(* IEC 61131-3 sources: traffic-lights/PLC_TrafficLights/Class/HwControl (part 2) *)

      ret_code                := BUSY;

      StartTime               := ops.tAbsolute;
      AdditionalPostInitTime  := 0;
      sd_retval               := 0;

//**********************************************************************************************************************************************************
//** CALCULATE, SET AND DISTRIBUTE TASK TIMES                                                                                                             **
//**********************************************************************************************************************************************************

      for i:=0 to TASK_SELECT_COREMAX do

      //Calculate Tasksettings for each core
        CalculateTaskInfo(us_CoreSelect:=i$USINT, pTaskInfo:=#aTaskInfoCore[i]);

        //Special Core 0 has to be running in RtWork method (is needed because if we dont have the new interfaces we cannot move a function to first realtime pos later)
        //Always add Realtime and Cyclic for Core 0: Realtime of Core 0 does watchdog trigger and calls for Diasmaster
        //***********************************************************
        if aTaskInfoCore[i].us_CoreSelect = TASK_SELECT_CORE0 then

          //Rt Prescan
          //**********************************************************************************************************************************************

          //get objectinfo of HwControl object
          //maybe we have a derivation with configured realtime task --> we have to change the task time of the task to the correct setting
          sd_retval := To_TaskObjectControl.GetObjectInfo( thispointer := this, tasktype := OBJ_RT, objinfo := #s_objinfo);

          //Check if we have a configured tasktime
          if sd_retval <> 0 | s_objinfo.period = 0 then

            //No task configured --> use OS function to add the RT Task

            //Note: udPhase must always be TASK_SCAN. At RTK there was an error that using TASK_PRE and TASK_POST occurs an access-exception in the OS.
            //With TASK_SCAN the object/function will be added in the list at the end. (will be moved to first position later if needed)
            if OS_AddRtObject(udMode  := TASK_TIMED
                            , udTime  := aTaskInfoCore[i].ud_MyRtTaskTime_us OR 16#8000_0000
                            , udPhase := TASK_SCAN) = NIL then
              HWC_LogValue1(this,"@0160 (HWControl::Control::NewInst) OS_AddRtObject failed to add Realtime (Prescan) object for core 0x{0}",aTaskInfoCore[i].us_CoreSelect);
            end_if;
          else

            // User must have a derivation of the HWControl with a configured Realtime Task --> Change the task time of the existing realtime task
            if To_TaskObjectControl.ChangeObjectState(thispointer :=  this
                                                    , actioncmd   :=  ACTION_NEWTIME
                                                    , tasktype    :=  OBJ_RT
                                                    , debugobj    :=  0
                                                    , newtime     :=  aTaskInfoCore[i].ud_MyRtTaskTime_us OR 16#8000_0000
                                                    ) <> 0 then
              HWC_LogError(this,"@03E3 (HWControl::Control::NewInst) Failed to change the object state to set the correct realtime task settings.");
            end_if;
          end_if;

          //RT Postscan
          //**********************************************************************************************************************************************

          //Check for Rt-Debug State. Do not add the Rt func for postscan if RtDebug is activated (because postscan will be called from prescan in this case)

          if GetRtDebugState() = TRUE then
            //save thispointer of object in OS-function (leads to that the task is called from the Breakpoint handler from the OS so the user can debug and the Hwcontrol is still running (no watchdog error))
            if p_DebugAPI then
              SaveThisPointer( this, TASK_SELECT_CORE0 );
            else
              HWC_LogError(this,"@0167 (HWControl::Control::NewInst) Pointer p_DebugAPI is invalid. Rt-Debug is not supported");
            end_if;

            // Set RtPostScan off if RtDebug is used!
            if To_TaskObjectControl.ChangeObjectState(thispointer :=  #HWRtPostScan.ClassSvr$void
                                                    , actioncmd   :=  ACTION_SUSPEND
                                                    , tasktype    :=  OBJ_RT
                                                    , debugobj    :=  0
                                                    , newtime     :=  0
                                                    ) <> 0 then
              HWC_LogError(this,"@0161 (HWControl::Control::NewInst) Failed to change object state of HwRtPostscan object");
            end_if;

          else

            //We have to use the object of HwRtPostscan instead of using the function OS_AddRtObject due to problems with RTK-CPUs (e.g. CP212)
            //The problem is that, with a maintimer of 500µs, and a task time of 1ms it can happen that the realtime (prescan) and the postscan of this class
            //are not "synchronized", which means that they have a time gap of 500µs between each other which leads to problems (TimesliceError).
            //This is not a problem with Salamander CPUs (e.g CP111)

            // Synchronize calls of Rt & RtPostScan (same timebase)
            if To_TaskObjectControl.ChangeObjectState(thispointer :=  #HWRtPostScan.ClassSvr$void
                                                    , actioncmd   :=  ACTION_NEWTIME
                                                    , tasktype    :=  OBJ_RT
                                                    , debugobj    :=  0
                                                    , newtime     :=  aTaskInfoCore[i].ud_MyRtTaskTime_us OR 16#8000_0000
                                                    ) <> 0 then
              HWC_LogError(this,"@0161 (HWControl::Control::NewInst) Failed to change object state of HwRtPostscan object");
            end_if;

            //save NIL-Pointer to OS-function because only HwControl is allowed to use this function
            if p_DebugAPI then
              SaveThisPointer( NIL, TASK_SELECT_CORE0 );
            end_if;

            //rt-post scan is added - realtime is added
            sRtTaskControl.usCoresRtActive  += 1;

          end_if;

          //Cyclic Task
          //**********************************************************************************************************************************************

          //Note: OS_AddCyFunc can NOT be used!! On RTK-CPUs with emulated SRAM () it leads to a reboot of the CPU if the SRAM is accessed from a function that is added via OS_AddCyFunc (or OS_AddRtFunc).
//          if OS_AddCyFunc (CyWork_CoreX
//                         , pParam  := #aTaskInfoCore[i].us_CoreSelect
//                         , udMode  := TASK_TIMED
//                         , udTime  := aTaskInfoCore[i].ud_MyCyTaskTime_us OR 16#8000_0000  //Time in µs instead of ms
//                         , udPhase := TASK_SCAN
//                          ) = NIL then
//
//            HWC_LogValue1(this,"@0162 (HWControl::Control::NewInst) OS_AddCyFunc failed to add Cyclic function for core 0x{0}",aTaskInfoCore[i].us_CoreSelect);
//          end_if;

          //get objectinfo of HwControl object
          //maybe we have a derivation with configured cyclic task --> we have to change the task time of the task to the correct setting
          sd_retval := To_TaskObjectControl.GetObjectInfo( thispointer := this, tasktype := OBJ_CT, objinfo := #s_objinfo );

          //Check if we have a configured tasktime
          if sd_retval <> 0 | s_objinfo.period = 0 then
            //No task configured --> use OS function to add the CY Task

            //Note: udPhase must always be TASK_SCAN. At RTK there was an error that using TASK_PRE and TASK_POST occurs an access-exception in the OS.
            //With TASK_SCAN the object/function will be added in the list at the end. (will be moved to first position later if needed)
            if OS_AddCyObject(udMode  := TASK_TIMED
                            , udTime  := aTaskInfoCore[i].ud_MyCyTaskTime_us OR 16#8000_0000
                            , udPhase := TASK_SCAN) = NIL then
              HWC_LogValue1(this,"@0160 (HWControl::Control::NewInst) OS_AddCyObject failed to add Cyclic object for core 0x{0}",aTaskInfoCore[i].us_CoreSelect);
            end_if;
          else

            // User must have a derivation of the HWControl with a configured cyclic Task --> Change the task time of the existing cyclic task
            if To_TaskObjectControl.ChangeObjectState(thispointer :=  this
                                                    , actioncmd   :=  ACTION_NEWTIME
                                                    , tasktype    :=  OBJ_CT
                                                    , debugobj    :=  0
                                                    , newtime     :=  aTaskInfoCore[i].ud_MyCyTaskTime_us OR 16#8000_0000
                                                    ) <> 0 then
              HWC_LogError(this,"@03E4 (HWControl::Control::NewInst) Failed to change the object state to set the correct cyclic task settings.");
            end_if;
          end_if;

        else

          //Check if core is needed
          if aTaskInfoCore[i].ud_MyRtTaskTime_us <> 0
           & aTaskInfoCore[i].ud_MyCyTaskTime_us <> 0 then

            //Check if new interfaces are available
            if Get_ITASK_Version() >= LSL_ITASK_VERSION_MULTICORE_SUPPORT then
              //Rt Prescan
              //**********************************************************************************************************************************************
#ifdef OS_AddRtFuncEx

              //Check if function pointer is valid. These function will never be valid on a RTK CPU because they don't support multicore features.
              //But maybe the ITASK Version will be extended for an other feature, so we will have an ITASK Version >= LSL_ITASK_VERSION_MULTICORE_SUPPORT at RTK CPUs
              if _LSL_POS^.piTask^.AddRealTimeFunctionEx <> NIL then

                if OS_AddRtFuncEx(RtPreScan_CoreX
                                , pParam  := #aTaskInfoCore[i].us_CoreSelect
                                , udMode  := TASK_TIMED
                                , udTime  := aTaskInfoCore[i].ud_MyRtTaskTime_us OR 16#8000_0000  //Time in µs instead of ms
                                , udPhase := TASK_SCAN
                                , core    := aTaskInfoCore[i].us_CoreSelect
                                ) = NIL then

                  HWC_LogValue1(this,"@0163 (HWControl::Control::NewInst) OS_AddRtFuncEx Failed to add Realtime (Prescan) function for core 0x{0}",aTaskInfoCore[i].us_CoreSelect);
                end_if;

                //Check if Rt-Debug is used
                if GetRtDebugState() = TRUE then

                  //Check if the new function is supported by the OS
                  if p_DebugAPI & p_DebugAPI^.version >= DEBUG_API_VERSION_MULTICORE_SUPPORT then
#ifdef SaveFunction
                    //Check if pointer is valid
                    if p_DebugAPI^.pSaveFunction <> NIL then
                      SaveFunction(#RtPreScan_CoreX(), this, aTaskInfoCore[i].us_CoreSelect);
                    else
                      HWC_LogError(this,"@0164 (HWControl::Control::NewInst) p_DebugAPI^.SaveFunction is nil. Rt-Debug is not supported.");
                    end_if;

#else
                    HWC_LogError(this,"@0165 (HWControl::Control::NewInst) Rt-Debug for multicore is not supported. SaveFunction is not defined.");
#endif
                  elsif p_DebugAPI then
                    HWC_LogError(this,"@0166 (HWControl::Control::NewInst) RT-Debug for multicore is not supported with this OS.");
                  else
                    HWC_LogError(this,"@0167 (HWControl::Control::NewInst) Pointer p_DebugAPI is invalid. Rt-Debug is not supported");
                  end_if;
                else
                  if p_DebugAPI & p_DebugAPI^.version >= DEBUG_API_VERSION_MULTICORE_SUPPORT then
#ifdef SaveFunction
                    if p_DebugAPI^.pSaveFunction <> NIL then
                      SaveFunction(#RtPreScan_CoreX(), nil, aTaskInfoCore[i].us_CoreSelect);
                    end_if;
#endif
                  elsif p_DebugAPI then
                    HWC_LogError(this,"@0166 (HWControl::Control::NewInst) RT-Debug for multicore is not supported with this OS.");
                  else
                    HWC_LogError(this,"@0167 (HWControl::Control::NewInst) Pointer p_DebugAPI is invalid. Rt-Debug is not supported");
                  end_if;
                end_if;

              else
                HWC_LogError(this,"@0168 (HWControl::Control::NewInst) Function pointer of _LSL_POS^.piTask^.AddRealTimeFunctionEx is invalid.");
              end_if;
#else
              //Log that function is not supported by Lasal
              //Only log here once
              HWC_LogError(this,"@0169 (HWControl::Control::NewInst) Warning! Unsupported LASAL-Class2 version detected to use OS_AddRtFuncEx function. Version 02.02.172 or higher is required to use this function");
#endif

              //RT Postscan
              //**********************************************************************************************************************************************
#ifdef OS_AddRtFuncEx
              //Check if function pointer is valid. These function will never be valid on a RTK CPU because they don't support multicore features.
              //But maybe the ITASK Version will be extended for an other feature, so we will have an ITASK Version >= LSL_ITASK_VERSION_MULTICORE_SUPPORT at RTK CPUs
              if _LSL_POS^.piTask^.AddRealTimeFunctionEx <> NIL then

                //Don't start Rt Postscan if RT-Debug is used (PostscanWork will be called from Prescan)
                if GetRtDebugState() = FALSE then

                  if OS_AddRtFuncEx(RtPostScan_CoreX
                                  , pParam  := #aTaskInfoCore[i].us_CoreSelect
                                  , udMode  := TASK_TIMED
                                  , udTime  := aTaskInfoCore[i].ud_MyRtTaskTime_us OR 16#8000_0000  //Time in µs instead of ms
                                  , udPhase := TASK_SCAN
                                  , core    := aTaskInfoCore[i].us_CoreSelect
                                  ) = NIL then

                    HWC_LogValue1(this,"@016A (HWControl::Control::NewInst) OS_AddRtFuncEx failed to add Realtime (Postscan) function for core 0x{0}",aTaskInfoCore[i].us_CoreSelect);
                  else
                    //rt-post scan is added - realtime is added
                    sRtTaskControl.usCoresRtActive  += 1;
                  end_if;
                else
                  HWC_LogError(this, "@016B (HWControl::Control::NewInst) RtDebug is used - RtPostScan is not possible together with RtDebug!");
                end_if;
              else
                HWC_LogError(this,"@0168 (HWControl::Control::NewInst) Function pointer of _LSL_POS^.piTask^.AddRealTimeFunctionEx is invalid.");
              end_if;
#endif

              //Cyclic Task
              //**********************************************************************************************************************************************
#ifdef OS_AddCyFuncEx

              //Check if function pointer is valid. These function will never be valid on a RTK CPU because they don't support multicore features.
              //But maybe the ITASK Version will be extended for an other feature, so we will have an ITASK Version >= LSL_ITASK_VERSION_MULTICORE_SUPPORT at RTK CPUs
              if _LSL_POS^.piTask^.AddCyclicFunctionEx <> NIL then

                if OS_AddCyFuncEx(CyWork_CoreX
                                , pParam  := #aTaskInfoCore[i].us_CoreSelect
                                , udMode  := TASK_TIMED
                                , udTime  := aTaskInfoCore[i].ud_MyCyTaskTime_us OR 16#8000_0000  //Time in µs instead of ms
                                , udPhase := TASK_SCAN
                                , core    := aTaskInfoCore[i].us_CoreSelect
                                ) = NIL then

                  HWC_LogValue1(this,"@016C (HWControl::Control::NewInst) OS_AddCyFuncEx failed to add Cyclic function for core 0x{0}",aTaskInfoCore[i].us_CoreSelect);
                end_if;
              else
                HWC_LogError(this,"@016D (HWControl::Control::NewInst) Function pointer of _LSL_POS^.piTask^.AddCyclicFunctionEx is invalid.");
              end_if;
#endif
            end_if;
          end_if;
        end_if;
      end_for;

      //read client setting for task synchronization
      RtTaskSync := RtTaskSync.Read() <> 0;

      if RtTaskSync = 1 then
        //check if more than one core is active and more than one rt task is available
        if sRtTaskControl.usCoresRtActive > 1 & ud_CPUCoreCount > 1 & us_CPUsRtCyEnabled > 1 then
          //search for different task times
          for i := 1 to sRtTaskControl.usCoresRtActive-1 do
            if aTaskInfoCore[0].ud_MyRtTaskTime_us <> aTaskInfoCore[i].ud_MyRtTaskTime_us then
              //task times are different - synchronizing is not possible
              RtTaskSync := 0;
              HWC_LogError(this, "@06AC (HwControl::Control::NewInst) The Rt task times are different so synchronization is not possible!");
              exit;
            end_if;
          end_for;

          if (mt_api = nil) & RtTaskSync = 1 then
            if(OS_CILGet("LSL_MULTITASK", #mt_api$void)) THEN
              mt_api := NIL;
              HWC_LogError(this,"@06AD (HWControl::Control::NewInst) Pointer for event semaphore is invalid. Synchronizing of Rt tasks is not supported!");
            else
              sRtTaskControl.pvPreRtSyncTaskEvent := OS_MT_CreateSemaphore(MTSEMATYPE_EVENT, 0, 0, "HwControl_PreRtSyncTaskEvent");
              sRtTaskControl.pvPostRtSyncTaskEvent := OS_MT_CreateSemaphore(MTSEMATYPE_EVENT, 0, 0, "HwControl_PostRtSyncTaskEvent");
              if sRtTaskControl.pvPreRtSyncTaskEvent <> NIL & sRtTaskControl.pvPostRtSyncTaskEvent <> NIL then
                //activate rt task synchronizing
                sRtTaskControl.b_RtTaskControlActive := TRUE;
              else
                //adding event semaphore for synchronizing task doesn't work
                HWC_LogError(this,"@06AF (HWControl::Control::NewInst) Pointer for event semaphore is invalid. Synchronizing of Rt tasks is not supported!");
              end_if;
            end_if;
          end_if;
        else
          HWC_LogError(this,"@06B0 (HWControl::Control::NewInst) There is only one Rt task available! Synchronizing of Rt tasks is deactivated.");
        end_if;
      end_if;

      //set client to actual setting
      RtTaskSync := sRtTaskControl.b_RtTaskControlActive;

      //Set Varanmanager variables (was done in AddVaranManager before, now we have to set these here because we know the task times just yet)
      //**************************************************************************

      //Go through all varanmanagers
      pOneManager := #a_VaranManager[0];

      for i := 0 to ( MAX_VARAN_MANAGERS - 1 ) do
        for j:= 0 to TASK_SELECT_COREMAX  do
          //Check if manager is available, set for right core and has set a time
          if ( pOneManager^.p_Functions         <> NIL
             & pOneManager^.p_Functions^.p_This <> NIL
             & pOneManager^.us_CoreSelect     = j
             )
          then
            pOneManager^.ud_SuperiorSync       := (pOneManager^.p_Functions^.ud_SuperiorTime / 1000 ) / (aTaskInfoCore[j].ud_MyRtTaskTime_us);
            pOneManager^.ud_SuperiorSyncActual := pOneManager^.ud_SuperiorSync;

      //       if the own tasktime is slower then superior varantime, don't wait for HW-Class Synchronity
            if (aTaskInfoCore[j].ud_MyRtTaskTime_us) > (pOneManager^.p_Functions^.ud_SuperiorTime / 1000) then
              pOneManager^.p_Functions^.b_HWClassSynchron    := TRUE;
              pOneManager^.p_Functions^.b_OverrideFrameCheck := TRUE;
            end_if;
          end_if;
        end_for;
        pOneManager += sizeof(t_OneVaranManager);
      end_for;

      //Distribute Task times to all connected classes
      //**************************************************************************
      MyPara.uiCmd := CMD_POST_INIT_DISTRIBUTE_TASKTIMES;

      MyPara.aPara[0]$t_Distribute_TaskTimes_Cmd.udVersion := 1;  //Version of command

      for i:=0 to TASK_SELECT_COREMAX do

        MyPara.aPara[0]$t_Distribute_TaskTimes_Cmd.udRtTaskTime_us := aTaskInfoCore[i].ud_MyRtTaskTime_us;  //Realtime Task time in µs
        MyPara.aPara[0]$t_Distribute_TaskTimes_Cmd.udCyTaskTime_us := aTaskInfoCore[i].ud_MyCyTaskTime_us;  //Cyclic Task time in µs

        //Check if task is active/needed
        if aTaskInfoCore[i].ud_MyRtTaskTime_us <> 0 & aTaskInfoCore[i].ud_MyCyTaskTime_us <> 0 then

          //We don't need to distribute the info to the Varanmanagers because the HwControl handles the time sheduling of the managers
          //Neither we distribute the info to the special objects

          // objects, which are controlled by HwControl (BusInterfaceSDIASInternal, Safetymanager,...)
          if pHwControlLogins then
            pHelp := pHwControlLogins;
            while pHelp <> NIL do
              // Check if its the right core
              if pHelp^.us_CoreSelect = i then
                pHelp^.pThis^.NewInst(pPara:=#MyPara, pResult:=#MyResult);
              end_if;
              pHelp := pHelp^.pNext;
            end_while;
          end_if;

          //First-Call Objects
          if pCallFirstObjects then
            pHelpFirst := pCallFirstObjects;
            while pHelpFirst <> NIL do
              // Check if its the right core
              if pHelpFirst^.us_CoreSelect = i then
                pHelpFirst^.pThis^.NewInst(pPara:=#MyPara, pResult:=#MyResult);
              end_if;
              pHelpFirst := pHelpFirst^.pNext;
            end_while;
          end_if;

        end_if;
      end_for;

//**********************************************************************************************************************************************************
//** INITIALIZE EVERYTHING VIA ASYNCHRON ACCESSES                                                                                                         **
//**********************************************************************************************************************************************************

      while (ret_code = BUSY) do
        // check the varanmanagers if they are not ready
        ret_code := READY;

        // only if there is a varan manager
        if VaranManagersAvailable then
          //call the last init of all varan managers
          pOneManager := #a_VaranManager[0];  // RamAnd: using pointers instead of array accesses reduces compiled awl-code by 120 lines!!!
          for i := 0 to ( MAX_VARAN_MANAGERS - 1 ) do

            //look if we have a correct pointer
            if ( pOneManager^.p_Functions & pOneManager^.p_Functions^.p_This ) then
              TempRetCode := pOneManager^.p_Functions^.p_This^.NewInst(pPara, pResult);

              // if any manager is still busy, we have to keep calling them
              if TempRetCode = BUSY then
                ret_code := TempRetCode;
              end_if;
            end_if;

            pOneManager += sizeof(t_OneVaranManager);
          end_for;
        end_if;

        // objects, which are controlled by HwControl
        if pHwControlLogins then
          pHelp := pHwControlLogins;
          while pHelp <> NIL do
            if pHelp^.bdSettings.PostInit then
              TempRetCode := pHelp^.pThis^.NewInst(pPara, pResult);
              // if any manager is still busy, we have to keep calling them
              if TempRetCode = BUSY then
                ret_code := TempRetCode;
              end_if;
            end_if;

            pHelp := pHelp^.pNext;
          end_while;
        end_if;

        // check timeout
        if ((ops.tAbsolute - StartTime) > (POST_INIT_TIMEOUT + AdditionalPostInitTime)) then
          HWC_LogError(this, "@016E (HwControl::Control::NewInst) Timeout in PostInit (initialize)");

          // only if there is a varan manager
          if VaranManagersAvailable then

            // Force all VM to end the PostInit Phase, Otherwise UpdateCy of HWK will not be called -----------------------------------------
            MyPara.uiCmd := CMD_FORCE_POST_INIT_END;

            //call the last init of all varan managers
            pOneManager := #a_VaranManager[0];
            for i := 0 to ( MAX_VARAN_MANAGERS - 1 ) do

              //look if we have a correct pointer
              if ( pOneManager^.p_Functions & pOneManager^.p_Functions^.p_This ) then
                TempRetCode := pOneManager^.p_Functions^.p_This^.NewInst(#MyPara, #MyResult);
              end_if;

              pOneManager += sizeof(t_OneVaranManager);
            end_for;	// ---------------------------------------------------------------------------------------------------------------------------------------------
          end_if;
          exit;
        end_if;
      end_while;

//**********************************************************************************************************************************************************
//** SORT THE VARAN DOs NEEDED FOR SAFETY                                                                                                                 **
//**********************************************************************************************************************************************************

      MyPara.uiCmd := CMD_POST_INIT_DO_SORT;

      // only if there is a varan manager
      if VaranManagersAvailable then
        //send the finish command to all varan managers
        pOneManager := #a_VaranManager[0];
        for i := 0 to ( MAX_VARAN_MANAGERS - 1 ) do

          //look if we have a correct pointer
          if ( pOneManager^.p_Functions & pOneManager^.p_Functions^.p_This ) then
            TempRetCode := pOneManager^.p_Functions^.p_This^.NewInst(pPara:=#MyPara, pResult:=#MyResult);

            // if any manager is still busy, we have to keep calling them
            if TempRetCode = BUSY then
              ret_code := TempRetCode;
            end_if;
          end_if;

          pOneManager += sizeof(t_OneVaranManager);
        end_for;
      end_if;

//**********************************************************************************************************************************************************
//** START THE REALTIME OF HWCONTROL                                                                                                                      **
//**********************************************************************************************************************************************************

      //bring HwControl to the first realtime task position and start realtime task

      //Check if the new LSL_ITASK functions are supported from the OS
      if Get_ITASK_Version() >= LSL_ITASK_VERSION_MULTICORE_SUPPORT then

        for i:= 0 to TASK_SELECT_COREMAX do

          //Special case for Realtime of Core 0 because it has the Standard RTWork Function
          if aTaskInfoCore[i].us_CoreSelect = TASK_SELECT_CORE0 then

            //Use the old (non multicore/extended) functions for Core 0 (Old OS will support this interface)
            OS_MoveObject(thisPtr   := this
                        , tasktype  := TASK_OBJ_RT
                        , flags     := 1 );

            OS_SetNbrOfLdrPhaseObjects(nbrOfObjs := 1);

          // Check if we have time settings for the current core
          elsif aTaskInfoCore[i].ud_MyRtTaskTime_us <> 0 & aTaskInfoCore[i].ud_MyCyTaskTime_us <> 0 then

#ifdef OS_MoveFunctionEx
            //Check if function pointer is valid. These function will never be valid on a RTK CPU because they don't support multicore features.
            //But maybe the ITASK Version will be extended for an other feature, so we will have an ITASK Version >= LSL_ITASK_VERSION_MULTICORE_SUPPORT at RTK CPUs
            if _LSL_POS^.piTask^.MoveFunctionEx <> NIL then

              //Move RtPreScan function to the first realtime task position of the selected core
              sd_retval := OS_MoveFunctionEx(pFunc     := #RtPreScan_CoreX()
                                           , pParam    := #aTaskInfoCore[i].us_CoreSelect
                                           , taskType  := TASK_OBJ_RT
                                           , flags     := 1
                                           , core      := aTaskInfoCore[i].us_CoreSelect);

              if sd_retval <> 0 then
                HWC_LogValue1(this,"@016F (HWControl::Control::NewInst) Function OS_MoveFunctionEx failed with retcode 0x{0}.", sd_retval$UDINT);
              end_if;
            else
              HWC_LogError(this,"@0170 (HWControl::Control::NewInst) Function pointer of _LSL_POS^.piTask^.MoveFunctionEx is invalid.");
            end_if;
#endif

#ifdef OS_SetNbrOfLdrPhaseObjectsEx

            //Check if function pointer is valid. These function will never be valid on a RTK CPU because they don't support multicore features.
            //But maybe the ITASK Version will be extended for an other feature, so we will have an ITASK Version >= LSL_ITASK_VERSION_MULTICORE_SUPPORT at RTK CPUs
            if _LSL_POS^.piTask^.SetNbrOfLdrPhaseObjectsEx <> NIL then

              sd_retval := OS_SetNbrOfLdrPhaseObjectsEx(nbrOfObjs := 1, core := aTaskInfoCore[i].us_CoreSelect);

              if sd_retval <> 0 then
                HWC_LogValue1(this,"@0171 (HWControl::Control::NewInst) Function OS_SetNbrOfLdrPhaseObjectsEx failed with retcode 0x{0}.", sd_retval$UDINT);
              end_if;

            else
              HWC_LogError(this,"@0172 (HWControl::Control::NewInst) Function pointer of _LSL_POS^.piTask^.SetNbrOfLdrPhaseObjectsEx is invalid.");
            end_if;

#endif
          end_if;
        end_for;

      else
        //Old version, multicore not supported, just bring realtime of core 0 to first position and start it
        OS_MoveObject(thisPtr   := this
                    , tasktype  := TASK_OBJ_RT
                    , flags     := 1 );

        OS_SetNbrOfLdrPhaseObjects(nbrOfObjs := 1);
      end_if;

//**********************************************************************************************************************************************************
//** WAIT FOR RT TO TAKE OVER THE WATCHDOG TRIGGERING                                                                                                     **
//**********************************************************************************************************************************************************

      MyPara.uiCmd            := CMD_POST_INIT_RT_SYNC;
      ret_code                := BUSY;

      StartTime               := ops.tAbsolute;
      AdditionalPostInitTime  := 0;

      while (ret_code = BUSY) do
        // check the varanmanagers if they are not ready
        ret_code := READY;

        // only if there is a varan manager
        if VaranManagersAvailable then
          //send the finish command to all varan managers
          pOneManager := #a_VaranManager[0];
          for i := 0 to ( MAX_VARAN_MANAGERS - 1 ) do

            //look if we have a correct pointer
            if ( pOneManager^.p_Functions & pOneManager^.p_Functions^.p_This ) then
              TempRetCode := pOneManager^.p_Functions^.p_This^.NewInst(pPara:=#MyPara, pResult:=#MyResult);

              // if any manager is still busy, we have to keep calling them
              if TempRetCode = BUSY then
                ret_code := TempRetCode;
              end_if;
            end_if;

            pOneManager += sizeof(t_OneVaranManager);
          end_for;
        end_if;

        // objects, which are controlled by HwControl
        if pHwControlLogins then
          pHelp := pHwControlLogins;
          while pHelp <> NIL do
            if pHelp^.bdSettings.PostInit then
              TempRetCode := pHelp^.pThis^.NewInst(pPara:=#MyPara, pResult:=#MyResult);
              // if any manager is still busy, we have to keep calling them
              if TempRetCode = BUSY then
                ret_code := TempRetCode;
              end_if;
            end_if;

            pHelp := pHelp^.pNext;
          end_while;
        end_if;

        // check timeout
        if ((ops.tAbsolute - StartTime) > (POST_INIT_TIMEOUT + AdditionalPostInitTime)) then
          HWC_LogError(this, "@0173 (HwControl::Control::NewInst) Timeout in PostInit (rt sync)");

          // only if there is a varan manager
          if VaranManagersAvailable then

            // Force all VM to end the PostInit Phase, Otherwise UpdateCy of HWK will not be called -----------------------------------------
            MyPara.uiCmd := CMD_FORCE_POST_INIT_END;

            //call the last init of all varan managers
            pOneManager := #a_VaranManager[0];  // RamAnd: using pointers instead of array accesses reduces compiled awl-code by 120 lines!!!
            for i := 0 to ( MAX_VARAN_MANAGERS - 1 ) do

              //look if we have a correct pointer
              if ( pOneManager^.p_Functions & pOneManager^.p_Functions^.p_This ) then
                TempRetCode := pOneManager^.p_Functions^.p_This^.NewInst(#MyPara, #MyResult);
              end_if;

              pOneManager += sizeof(t_OneVaranManager);
            end_for;	// ---------------------------------------------------------------------------------------------------------------------------------------------
          end_if;
          exit;
        end_if;
      end_while;

//**********************************************************************************************************************************************************
//** LOAD THE SAFETY PROJECT CONFIGURATIONS AT THE SAFETY CPUS                                                                                            **
//**********************************************************************************************************************************************************

      // tell the available safety cpu modules to get their configurations now!
      MyPara.uiCmd := CMD_SM_POST_INIT_FINISHED;
      SafetyManager.ClassState.NewInst(pPara:=#MyPara, pResult:=#MyResult);

//**********************************************************************************************************************************************************
//** FINISH DIAS/CDIAS                                                                                                                                    **
//**********************************************************************************************************************************************************

      //look if DiasMaster is also used ( must be after starting realtime task )
      if ( s_DiasMaster.p_Functions <> NIL ) then

        //make final initialization in DiasMaster
        CallPtr	( p_function	:= s_DiasMaster.p_Functions^.p_LastInit
                , p_this		  := s_DiasMaster.p_Functions^.p_This
                );
      end_if;

//**********************************************************************************************************************************************************
//** FINISH VARAN/SDIAS                                                                                                                                   **
//**********************************************************************************************************************************************************

      MyPara.uiCmd            := CMD_POST_INIT_RT_READY;
      ret_code                := BUSY;

      StartTime               := ops.tAbsolute;
      AdditionalPostInitTime  := 0;

      while (ret_code = BUSY) do
        // check the varanmanagers if they are not ready
        ret_code := READY;

        // only if there is a varan manager
        if VaranManagersAvailable then
          //send the finish command to all varan managers
          pOneManager := #a_VaranManager[0];
          for i := 0 to ( MAX_VARAN_MANAGERS - 1 ) do

            //look if we have a correct pointer
            if ( pOneManager^.p_Functions & pOneManager^.p_Functions^.p_This ) then
              TempRetCode := pOneManager^.p_Functions^.p_This^.NewInst(pPara:=#MyPara, pResult:=#MyResult);

              // if any manager is still busy, we have to keep calling them
              if TempRetCode = BUSY then
                ret_code := TempRetCode;
              end_if;
            end_if;

            pOneManager += sizeof(t_OneVaranManager);
          end_for;
        end_if;

        // objects, which are controlled by HwControl
        if pHwControlLogins then
          pHelp := pHwControlLogins;
          while pHelp <> NIL do
            if pHelp^.bdSettings.PostInit then
              TempRetCode := pHelp^.pThis^.NewInst(pPara:=#MyPara, pResult:=#MyResult);
              // if any manager is still busy, we have to keep calling them
              if TempRetCode = BUSY then
                ret_code := TempRetCode;
              end_if;
            end_if;

            pHelp := pHelp^.pNext;
          end_while;
        end_if;

        // check timeout
        if ((ops.tAbsolute - StartTime) > (POST_INIT_TIMEOUT + AdditionalPostInitTime)) then
          HWC_LogError(this, "@0174 (HwControl::Control::NewInst) Timeout in PostInit (finishing)");

          // only if there is a varan manager
          if VaranManagersAvailable then

            // Force all VM to end the PostInit Phase, Otherwise UpdateCy of HWK will not be called -----------------------------------------
            MyPara.uiCmd := CMD_FORCE_POST_INIT_END;

            //call the last init of all varan managers
            pOneManager := #a_VaranManager[0];  // RamAnd: using pointers instead of array accesses reduces compiled awl-code by 120 lines!!!
            for i := 0 to ( MAX_VARAN_MANAGERS - 1 ) do

              //look if we have a correct pointer
              if ( pOneManager^.p_Functions & pOneManager^.p_Functions^.p_This ) then
                TempRetCode := pOneManager^.p_Functions^.p_This^.NewInst(#MyPara, #MyResult);
              end_if;

              pOneManager += sizeof(t_OneVaranManager);
            end_for;	// ---------------------------------------------------------------------------------------------------------------------------------------------
          end_if;
          exit;
        end_if;
      end_while;

//**********************************************************************************************************************************************************
//** Tell everything that the Post-Init is Done                                                                                                           **
//**********************************************************************************************************************************************************

      // Tell DiasMaster that the Post-Init is Done
      // needed for CallRealtime_IM
      MyPara.uiCmd := CMD_SET_POSTINIT_DONE;

      if s_DiasMaster.p_Functions then
        ret_code := s_DiasMaster.p_Functions^.p_This$pVirtualBase^.NewInst(#MyPara, pResult:=#MyResult);
      end_if;

      // only if there is a varan manager
      if VaranManagersAvailable then
        //send the finish command to all varan managers
        pOneManager := #a_VaranManager[0];
        for i := 0 to ( MAX_VARAN_MANAGERS - 1 ) do

          //look if we have a correct pointer
          if ( pOneManager^.p_Functions & pOneManager^.p_Functions^.p_This ) then
            TempRetCode := pOneManager^.p_Functions^.p_This^.NewInst(pPara:=#MyPara, pResult:=#MyResult);

            // if any manager is still busy, we have to keep calling them
            if TempRetCode = BUSY then
              ret_code := TempRetCode;
            end_if;
          end_if;

          pOneManager += sizeof(t_OneVaranManager);
        end_for;
      end_if;

      // objects, which are controlled by HwControl
      if pHwControlLogins then
        pHelp := pHwControlLogins;
        while pHelp <> NIL do
          if pHelp^.bdSettings.PostInit then
            TempRetCode := pHelp^.pThis^.NewInst(pPara:=#MyPara, pResult:=#MyResult);
            // if any manager is still busy, we have to keep calling them
            if TempRetCode = BUSY then
              ret_code := TempRetCode;
            end_if;
          end_if;
          pHelp := pHelp^.pNext;
        end_while;
      end_if;

      bPostInitFinished := TRUE;  //Remember that post init is finished

#ifdef HWC_ENABLE_SPAM_PROTECTION
      // stop the override => from now on the spam protection is active
      HwcLogging.OverrideSpamProtection.Write(input:=0);
#endif

//**********************************************************************************************************************************************************
    CMD_GET_SUPPORTED_FEATURES:

      //Set length to be flexible for future
      pResult^.uiLng := 4;
      pResult^.aData[0]$BDINT := SupportedFeatures;

//**********************************************************************************************************************************************************
    CMD_HWCONTROL_LOGIN:
      TempSettings  := pPara^.aPara[1]$t_HwObjListSettings;
      us_ModuleType := pPara^.aPara[2]$USINT;
      us_CoreSelect := pPara^.aPara[3]$USINT;
      ud_RtTime_us  := pPara^.aPara[4]$UDINT;
      ud_CyTime_us  := pPara^.aPara[5]$UDINT;

      if (us_ModuleType AND HWT_ESCAPE_SEQU) = 0 then
        us_ModuleType := 0; // MSB must be set for a valid Escape Sequence
      end_if;

      if AddHwObject( pThis           :=  pPara^.aPara[0]$pVirtualBase
                    , Settings        :=  TempSettings
                    , EscapeSequence  :=  us_ModuleType
                    , us_CoreSelect   :=  us_CoreSelect
                    , ud_RtTime_us    :=  ud_RtTime_us
                    , ud_CyTime_us    :=  ud_CyTime_us
                    ) <> 0 then

        ret_code := ERROR;
      end_if;

      pResult^.uiLng          := 8;
      //Just return value of maintimer in ns to be compatible
      //Old classes --> do not set a new time --> task will be started with maintimer as time, so they will get the right time
      //New classes don't proove the return values, because the times will be distributed at the beginning of the post init phase
      pResult^.aData[0]$UDINT := _ClockTicks * 1000;
      pResult^.aData[4]$UDINT := _ClockTicks * 1000;

      // post init callback is only possible if the method is supported by loader
      if TempSettings.PostInit & (InstallPostInitCB() <> 0) then
        ret_code := ERROR;
      end_if;

//**********************************************************************************************************************************************************
  CMD_GET_HARDWARE_TREE_ENTRY:

    //Reset all Return Values
    pResult^.aData$t_HWCGetHardwareTreeEntryOut.pStr_NextHardewareTreeEntry := nil;
    pResult^.aData$t_HWCGetHardwareTreeEntryOut.retcode                     := _HWC_RETVAL_ERROR;
    ret_code                                                                := ERROR;

    pStr_HWTreeEntry  :=  pPara^.aPara[0]$t_HWCGetHardwareTreeEntryIn.pStr_LastHardewareTreeEntry;

    //Standard: Use varan manager number 0
    usVaranManagerNrTreeEntry := 0;

    // if nil, search the first module ==================================================================================================================
    if pPara^.aPara$t_HWCGetHardwareTreeEntryIn.pStr_LastHardewareTreeEntry = nil then

      // Call all managers and search the module
      us_ModuleType := HWT_ESCAPE_VARAN; // 1. entry requested, start with Varan HWKs

    //Search the next module =============================================================================================================================
    //Only when there is a valid length we can access the data
    elsif (pStr_HWTreeEntry$^UINT^ <> 0) then // Length is 2 byte

      // 3 byte is domain
      // 4 byte is bus type/escape sequence.
      us_ModuleType := (pStr_HWTreeEntry+3)^$USINT;

      //Current Index = 4 because first 2 bytes are length, one byte domain number, next byte is escape sequence, 5th byte is port number
      pPara^.aPara[0]$t_HWCGetHardwareTreeEntryIn.us_current_index  := 4;  //points to escape sequence

      //Current length is length - 2 (point above domain number and escape sequence)
      pPara^.aPara[0]$t_HWCGetHardwareTreeEntryIn.us_current_length$UINT := pStr_HWTreeEntry^$UINT - 2;

      //Multivaran-Manager Support:
      //Check if our module type is the multivaran escape sequence
      if us_ModuleType = HWT_ESCAPE_MULTIVARAN then
        us_ModuleType := (pStr_HWTreeEntry+5)^$USINT;

        //Get the varan manager number of the module
        usVaranManagerNrTreeEntry := (pStr_HWTreeEntry+4)^$USINT;

        //Increment index + 2 (ESCAPE-SEQUENZ MULTIVARAN + ManagerNumber)
        pPara^.aPara[0]$t_HWCGetHardwareTreeEntryIn.us_current_index  += 2;  //points to escape sequence

        //Increment length + 2(ESCAPE-SEQUENZ MULTIVARAN + ManagerNumber)
        pPara^.aPara[0]$t_HWCGetHardwareTreeEntryIn.us_current_length$UINT += 2;

      end_if;

    end_if;

    //Go through all managers

    //Varan -------------------------------------------------------------------------------------------------------------------
    if us_ModuleType = HWT_ESCAPE_VARAN then

      // Loop over all Varanmanger
      //Point to correct manager with the index
      pOneManager := #a_VaranManager[usVaranManagerNrTreeEntry];  // RamAnd: using pointers instead of array accesses reduces compiled awl-code by 120 lines!!!

      //look if we have a correct pointer
      if (pOneManager^.p_Functions) & ( pOneManager^.p_Functions^.p_This ) then
        ret_code := pOneManager^.p_Functions^.p_This^.NewInst(pPara, pResult);

        if (ret_code = READY) then

          if pResult^.aData[0]$t_HWCGetHardwareTreeEntryOut.retcode = _HWC_RETVAL_OK_HWTSTR_RETURNED then
            return; // Next HWT string was returned pass it back
          end_if;

          if pResult^.aData[0]$t_HWCGetHardwareTreeEntryOut.retcode = _HWC_RETVAL_OK_MODULE_FOUND |
             pResult^.aData[0]$t_HWCGetHardwareTreeEntryOut.retcode = _HWC_RETVAL_OK_END_OF_LIST then
            // Module was found and was the last module in the Manager
            // Set the requested HWT string to nil so that the next call is an autohit
            pPara^.aPara$t_HWCGetHardwareTreeEntryIn.pStr_LastHardewareTreeEntry := nil;

            ret_code := ERROR;  // Reset ret_code before next call

          end_if;

        end_if;

      end_if;

      // Try next Manager
      us_ModuleType := HWT_ESCAPE_CDIAS;
    end_if;

    //CDIAS DIAS -------------------------------------------------------------------------------------------------------------------
    if us_ModuleType = HWT_ESCAPE_CDIAS |
       us_ModuleType = HWT_ESCAPE_DIAS then

      if s_DiasMaster.p_Functions then

        ret_code := s_DiasMaster.p_Functions^.p_This$pVirtualBase^.NewInst(pPara,pResult);

        if pResult^.aData[0]$t_HWCGetHardwareTreeEntryOut.retcode = _HWC_RETVAL_OK_HWTSTR_RETURNED then
          return; // Next HWT string was returned pass it back
        end_if;

        if pResult^.aData[0]$t_HWCGetHardwareTreeEntryOut.retcode = _HWC_RETVAL_OK_MODULE_FOUND |
           pResult^.aData[0]$t_HWCGetHardwareTreeEntryOut.retcode = _HWC_RETVAL_OK_END_OF_LIST then
          // Module was found and was the last module in the Manager
          // Set the requested HWT string to nil so that the next call is an autohit
          pPara^.aPara$t_HWCGetHardwareTreeEntryIn.pStr_LastHardewareTreeEntry := nil;

          ret_code := ERROR;  // Reset ret_code before next call
        end_if;

      end_if;

      // Try next Manager
      us_ModuleType := HWT_ESCAPE_SEQU;

    end_if;

     // Other (Local SDIAS)  -------------------------------------------------------------------------------------------------------------------
    if us_ModuleType AND HWT_ESCAPE_SEQU then
      if pHwControlLogins then

        pHelp := pHwControlLogins;

        while pHelp <> NIL  do

          if pHelp^.usEscSequence AND HWT_ESCAPE_SEQU then

            ret_code := pHelp^.pThis^.NewInst(pPara, pResult);

            if pResult^.aData[0]$t_HWCGetHardwareTreeEntryOut.retcode = _HWC_RETVAL_OK_HWTSTR_RETURNED then
              return; // Next HWT string was returned pass it back
            end_if;

            if pResult^.aData[0]$t_HWCGetHardwareTreeEntryOut.retcode = _HWC_RETVAL_OK_MODULE_FOUND |
               pResult^.aData[0]$t_HWCGetHardwareTreeEntryOut.retcode = _HWC_RETVAL_OK_END_OF_LIST then
              // Module was found and was the last module in the Manager
              // Set the requested HWT string to nil so that the next call is an autohit
              pPara^.aPara$t_HWCGetHardwareTreeEntryIn.pStr_LastHardewareTreeEntry := nil;

              ret_code := ERROR;  // Reset ret_code before next call
            end_if;

          end_if;

          pHelp := pHelp^.pNext;

        end_while;

      end_if;

    end_if;

    // Check if no further module exits
    if pPara^.aPara$t_HWCGetHardwareTreeEntryIn.pStr_LastHardewareTreeEntry = nil then
      ret_code := READY;
      pResult^.aData[0]$t_HWCGetHardwareTreeEntryOut.retcode                      := _HWC_RETVAL_OK_END_OF_LIST;
      pResult^.aData[0]$t_HWCGetHardwareTreeEntryOut.pStr_NextHardewareTreeEntry  := NIL;

    end_if;

//**********************************************************************************************************************************************************
  CMD_GET_HARDWARE_DIAGNOSIS:

    pResult^.aData[0]$t_HWCGetHardwareDiagnosisOut.retcode := _HWC_RETVAL_ERROR;
    ret_code := ERROR;

    // Reset all return values
    pResult^.aData[0]$t_HWCGetHardwareDiagnosisOut.ClassState      := 16#FFFFFFFF$t_e_VaranErrors;  //invalid value
    pResult^.aData[0]$t_HWCGetHardwareDiagnosisOut.pStr_DeviceName := NIL;
    pResult^.aData[0]$t_HWCGetHardwareDiagnosisOut.ud_DeviceID     := HWC_INVALID_DEVICE_ID;
    pResult^.aData[0]$t_HWCGetHardwareDiagnosisOut.pStr_VendorName := NIL;
    pResult^.aData[0]$t_HWCGetHardwareDiagnosisOut.ud_VendorID     := 0;
    pResult^.aData[0]$t_HWCGetHardwareDiagnosisOut.pStr_SerialNo   := NIL;
    pResult^.aData[0]$t_HWCGetHardwareDiagnosisOut.pStr_OrderingNo := NIL;
    pResult^.aData[0]$t_HWCGetHardwareDiagnosisOut.ud_LicenseNo    := 0;
    pResult^.aData[0]$t_HWCGetHardwareDiagnosisOut.hd_HWVersion    := 0;
    pResult^.aData[0]$t_HWCGetHardwareDiagnosisOut.ud_Variante     := 0;
    pResult^.aData[0]$t_HWCGetHardwareDiagnosisOut.hd_FPGAVersion  := 0;
    pResult^.aData[0]$t_HWCGetHardwareDiagnosisOut.pStr_FWVersion  := NIL;
    pResult^.aData[0]$t_HWCGetHardwareDiagnosisOut.hd_SafetyNumber := 0;
    pResult^.aData[0]$t_HWCGetHardwareDiagnosisOut.ud_Place        := 16#FFFFFFFF; // Place 0 is valid
    pResult^.aData[0]$t_HWCGetHardwareDiagnosisOut.ud_AxisNo       := 16#FFFFFFFF;
    pResult^.aData[0]$t_HWCGetHardwareDiagnosisOut.ud_reserved_size:= 0;
    pResult^.aData[0]$t_HWCGetHardwareDiagnosisOut.pud_reserved    := NIL;
    pResult^.aData[0]$t_HWCGetHardwareDiagnosisOut.ud_user_size    := 0;
    pResult^.aData[0]$t_HWCGetHardwareDiagnosisOut.pud_user        := NIL;
    pResult^.aData[0]$t_HWCGetHardwareDiagnosisOut.p_DynExtList    := NIL;

    pStr_HWTRequested  :=  pPara^.aPara[0]$t_HWCGetHardwareDiagnosisIn.pStr_HardewareTreeEntry;

    //Only when there is a valid length we can access the data
    if (pStr_HWTRequested$^UINT^ <> 0) then // Length is 2 byte

      // 3 byte is domain

      // 4 byte is bus type/escape sequence.
      us_ModuleType := (pStr_HWTRequested+3)^$USINT;

      //Standard: Use varan manager number 0
      usVaranManagerNrTreeEntry := 0;

      //Current Index = 5 because first 2 bytes are length, one byte domain number, next byte is escape sequence, 5th byte is port number
      pPara^.aPara[0]$t_HWCGetHardwareDiagnosisIn.us_current_index  := 4;  //points to escape sequence
      //Current length is length - 2 (point above domain number and escape sequence)
      pPara^.aPara[0]$t_HWCGetHardwareDiagnosisIn.us_current_length$UINT := pStr_HWTRequested^$UINT - 2;

      //Multivaran-Manager Support:
      //Check if our module type is the multivaran escape sequence
      if us_ModuleType = HWT_ESCAPE_MULTIVARAN then

        us_ModuleType := (pStr_HWTRequested+5)^$USINT;

        //Get the varan manager number of the module
        usVaranManagerNrTreeEntry := (pStr_HWTRequested+4)^$USINT;

        //Increment index + 2 (ESCAPE-SEQUENZ MULTIVARAN + ManagerNumber)
        pPara^.aPara[0]$t_HWCGetHardwareTreeEntryIn.us_current_index  += 2;  //points to escape sequence

        //Increment length + 2(ESCAPE-SEQUENZ MULTIVARAN + ManagerNumber)
        pPara^.aPara[0]$t_HWCGetHardwareTreeEntryIn.us_current_length$UINT += 2;

      end_if;

      case us_ModuleType of

        //-------------------------------------------------------------------------------------------
        HWT_ESCAPE_VARAN:

          // Loop over all Varanmanger
          pOneManager := #a_VaranManager[usVaranManagerNrTreeEntry];  // RamAnd: using pointers instead of array accesses reduces compiled awl-code by 120 lines!!!

          //look if we have a correct pointer
          if (pOneManager^.p_Functions) & ( pOneManager^.p_Functions^.p_This ) then
            ret_code := pOneManager^.p_Functions^.p_This^.NewInst(pPara, pResult);
          end_if;

        //-------------------------------------------------------------------------------------------
        HWT_ESCAPE_CDIAS:

          if s_DiasMaster.p_Functions then
            ret_code := s_DiasMaster.p_Functions^.p_This$pVirtualBase^.NewInst(pPara,pResult);
          end_if;

        //-------------------------------------------------------------------------------------------
        HWT_ESCAPE_DIAS:

          if s_DiasMaster.p_Functions then
            ret_code := s_DiasMaster.p_Functions^.p_This$pVirtualBase^.NewInst(pPara,pResult);
          end_if;

        //-------------------------------------------------------------------------------------------
//        HWT_ESCAPE_SDIAS:

        // Other (SDIAS)
        else
          if pHwControlLogins then

            pHelp := pHwControlLogins;

            while pHelp <> NIL &
              ((ret_code <> READY) & (ret_code <> BUSY)) do // Module was found if retcode is ready or busy

              if pHelp^.usEscSequence = us_ModuleType then
                ret_code := pHelp^.pThis^.NewInst(pPara, pResult);
              end_if;

              pHelp := pHelp^.pNext;

            end_while;

          end_if;

      end_case;
    end_if;

//**********************************************************************************************************************************************************
  CMD_SET_VARANMANAGER_ERROR:

    //Raise manage error at all varan managers
    pOneManager := #a_VaranManager[0];
    for i := 0 to ( MAX_VARAN_MANAGERS - 1 ) do

      //look if we have a correct pointer
      if (pOneManager^.p_Functions) & ( pOneManager^.p_Functions^.p_This ) then
        pOneManager^.p_Functions^.p_This^.RaiseManagerError(pPara^.aPara[0]$UDINT);

      end_if;
      pOneManager += sizeof(t_OneVaranManager);
    end_for;

//**********************************************************************************************************************************************************
  CMD_EXTEND_POST_INIT_TIME:

    AdditionalPostInitTime += pPara^.aPara[0]$UDINT;

//**********************************************************************************************************************************************************
  CMD_LOGIN_VARANMANAGER:

    ret_code := READY;
    pResult^.aData[0]$DINT := AddVaranManager(ud_manager_number  := pPara^.aPara[0]$UDINT
                                            , p_function_list    := pPara^.aPara[1]$^void
                                            , us_CoreSelect      := pPara^.aPara[2]$USINT
                                            , ud_RtTime_us       := pPara^.aPara[3]$UDINT
                                            , ud_CyTime_us       := pPara^.aPara[4]$UDINT
                                            );

//**********************************************************************************************************************************************************
  CMD_DISABLE_VARANMANAGER:

    ret_code := READY;
    pResult^.aData[0]$DINT := DisableVaranManager(ud_manager_number := pPara^.aPara[0]$UDINT
                                                , p_function_list   := pPara^.aPara[1]$^void
                                                );

//**********************************************************************************************************************************************************
  CMD_GET_HW_TIMESTAMP:

    //NewInst CMD for SmartIO modules to fetch timestamp from HwControl

    ret_code := ERROR;

    // Version 1 does not support core select
    if pPara^.aPara[0]$t_GetHwTimestampCmd.udVersion = 1 then

      ret_code := READY;

      pResult^.uiLng      := sizeof(t_GetHwTimestampResult);
      pResult^.aData[0]$t_GetHwTimestampResult.udVersion   := 1;
      pResult^.aData[0]$t_GetHwTimestampResult.uiTimeStamp := aTaskInfoCore[TASK_SELECT_CORE0].uiHwTimeStamp_us;

    // Version 2 supports core selection
    elsif pPara^.aPara[0]$t_GetHwTimestampCmd.udVersion = 2 then

      ret_code := READY;
      us_CoreSelect := pPara^.aPara[0]$t_GetHwTimestampCmd.udCoreSelect$USINT;

      pResult^.uiLng      := sizeof(t_GetHwTimestampResult);
      pResult^.aData[0]$t_GetHwTimestampResult.udVersion   := 1;
      pResult^.aData[0]$t_GetHwTimestampResult.uiTimeStamp := aTaskInfoCore[us_CoreSelect].uiHwTimeStamp_us;

    end_if;
//**********************************************************************************************************************************************************

  CMD_HWC_REQ_PLLNS_REGULATION:

    ret_code := ERROR;

    //Version
    if pPara^.aPara[0] >= 1 then

      pResult^.uiLng := sizeof(DINT) + sizeof(t_HWCRetvalReturnCode);
      pResult^.aData[0]$DINT := 1;                 // Version

      if b_SoftwareSyncActive then
        pResult^.aData[4]   := _HWC_RETVAL_ERROR_SYNCREG_INUSE;//request denied  Software Synchronisation is already in use.
      else
        pResult^.aData[4]$t_HWCRetvalReturnCode := _HWC_RETVAL_OK;//request granted
        b_SoftwareSyncActive := TRUE;
      end_if;

      ret_code := READY;

    end_if;

    //**********************************************************************************************************************************************************

    //**********************************************************************************************************************************************************
    CMD_HWC_CONVERT_COMPRESSED_HWPATH:

      //Forward newinst to safety manager
      ret_code := SafetyManager.ClassState.NewInst(pPara:=pPara, pResult:=pResult);

  end_case;

END_FUNCTION

FUNCTION HwControl::InstallPostInitCB
  VAR_OUTPUT
    sd_retval 	: DINT;
  END_VAR
  VAR
    pFunction   : ^void;
  END_VAR

  sd_retval := -1;

  if b_PostInitInstalled = TRUE then
    sd_retval := 0;   // Return OK
  else

    // tell the loader that we need a post init phase
    pFunction := _FindFctName("LDR_InstallPostInitCB");
    if ( pFunction <> NIL ) then
      pFunction $ LDR_InstallPostInitCB(pThis:=this, pCmdSvr:=(#this^.Control.pMeth)$^SvrChCmd, newInstCmd:=CMD_POST_INIT_CALL);

      b_PostInitInstalled := TRUE;
      sd_retval           := 0;

    end_if;
  end_if;

END_FUNCTION

FUNCTION GLOBAL HwControl::DisableVaranManager
  VAR_INPUT
    ud_manager_number 	: UDINT;
    p_function_list 	: ^void;
  END_VAR
  VAR_OUTPUT
    sd_retval 	: DINT;
  END_VAR

  // is class ok
  if ( State = _ClassOk ) then

    // check pointer of watchdog interface
    if pSCDW = NIL then

      //look if it is a correct VaranManager number
      if (( ud_manager_number >= 0 ) &
          ( ud_manager_number <= MAX_VARAN_MANAGERS - 1 )) then

        // is this number already in use
        if ( a_VaranManager[ ud_manager_number ].p_Functions <> NIL ) then

          a_VaranManager[ ud_manager_number ].p_Functions	:= NIL;
          VaranManagersAvailable -= 1;
          sd_retval := 0;

        else
          sd_retval := -1;
          HWC_LogError(this, "@0175 (HwControl::DisableVaranManager) Manager is not even used!");
        end_if;
      else
        sd_retval := -2;
        HWC_LogError(this, "@0176 (HwControl::DisableVaranManager) Wrong VaranManagerNumber!");
      end_if;
    else
      sd_retval := -3;
      HWC_LogError(this, "@0177 (HwControl::DisableVaranManager) Called too late, the Watchdog is already active!");
    end_if;
  else
    sd_retval := -4;
    HWC_LogError(this, "@0178 (HwControl::DisableVaranManager) Class state is not ok!");
  end_if;

END_FUNCTION

FUNCTION HwControl::UpdateRtVaranManager
  VAR_INPUT
    usActiveCore 	: USINT;
  END_VAR
  VAR
    i			: DINT;
    pOneManager : ^t_OneVaranManager;
  END_VAR

  //update realtime functions of all VaranManagers
  //*****************************************************************************
  pOneManager := #a_VaranManager[0];  // RamAnd: using pointers instead of array accesses reduces compiled awl-code by 120 lines!!!
  for i := 0 to ( MAX_VARAN_MANAGERS - 1 ) do

    //look if right core, or call all manager if only one core is available
    if ( pOneManager^.us_CoreSelect = usActiveCore) then

      //look if we have a correct pointer
      if ( pOneManager^.p_Functions$^INT <> NIL ) then

        // if VMC is used, then check if the framecounter has been increased => right time to call Varan HW-Classes
        if (pOneManager^.p_Functions^.b_IsAlsoClient & (pOneManager^.p_Functions^.b_OverrideFrameCheck = FALSE) &
            pOneManager^.p_Functions^.p_This^.FrameCounterChanged(#pOneManager^.usOldFrameCnt, #pOneManager^.usActFrameCnt)) then

          // maybe we got some phase shift
          if (pOneManager^.ud_SuperiorSyncActual <> pOneManager^.ud_SuperiorSync) &
             (pOneManager^.ud_SuperiorSyncActual MOD pOneManager^.ud_SuperiorSync) then

            pOneManager^.ud_SuperiorSyncActual := pOneManager^.ud_SuperiorSync;
            pOneManager^.ud_CounterRt := pOneManager^.ud_RtTime_us;

            pOneManager^.usSyncCheck := 0; // reset synchronity
          end_if;
        end_if;

        //if call time for varan manager is reached
        if ( pOneManager^.ud_CounterRt = pOneManager^.ud_RtTime_us ) then

          //reset task time counter
          pOneManager^.ud_CounterRt := 0;

          //call realtime methode of VaranMaster
          pOneManager^.p_Functions^.p_This^.RtWork( 0 );

          // if manager is also client and we are in superior task
          if (pOneManager^.p_Functions^.b_IsAlsoClient = 1) & (pOneManager^.p_Functions^.b_OverrideFrameCheck = FALSE) then
            if (pOneManager^.ud_SuperiorSyncActual MOD pOneManager^.ud_SuperiorSync) = 0 then
              pOneManager^.ud_SuperiorSyncActual := 0;

              pOneManager^.usSyncCheck := (pOneManager^.usSyncCheck SHL 1) OR (pOneManager^.usActFrameCnt <> pOneManager^.usOldFrameCnt);

              if (pOneManager^.usSyncCheck = 16#FF) then
                pOneManager^.p_Functions^.b_HWClassSynchron := TRUE;
              else
                pOneManager^.p_Functions^.b_HWClassSynchron := FALSE;
              end_if;
            elsif (pOneManager^.ud_SuperiorSyncActual > pOneManager^.ud_SuperiorSync) then
              pOneManager^.ud_SuperiorSyncActual := 0;
            end_if;
          end_if;
        else
          if (pOneManager^.p_Functions^.b_IsAlsoClient & (pOneManager^.p_Functions^.b_OverrideFrameCheck = FALSE) &
             (((pOneManager^.p_Functions^.ud_SuperiorTime / 1000 ) > pOneManager^.ud_RtTime_us) |
             (pOneManager^.ud_SuperiorSyncActual MOD pOneManager^.ud_SuperiorSync)) &
             pOneManager^.p_Functions^.p_This^.FrameCounterChanged(#pOneManager^.usOldFrameCnt, #pOneManager^.usActFrameCnt)) then
            //set task time counter to HwControl task time
            pOneManager^.ud_CounterRt := 0;
            pOneManager^.ud_SuperiorSyncActual := 0;
            pOneManager^.usSyncCheck := 0;  // reset synchronity
          end_if;
        end_if;

        // add task time to counter
        pOneManager^.ud_CounterRt += aTaskInfoCore[usActiveCore].ud_MyRtTaskTime_us;

        // increase cycle counter
        pOneManager^.ud_SuperiorSyncActual += 1;
      end_if;
    end_if;

    pOneManager += sizeof(t_OneVaranManager);
  end_for;

END_FUNCTION

FUNCTION HwControl::UpdateRtPostScanVaranManager
  VAR_INPUT
    usActiveCore 	: USINT;
  END_VAR
  VAR
    i			: DINT;
    pOneManager : ^t_OneVaranManager;
  END_VAR

  //Update Rt PostScan method of all varanmanagers
  //*****************************************************************************
  pOneManager := #a_VaranManager[0];
  for i := 0 TO (MAX_VARAN_MANAGERS - 1) do
    //Look for right core
    if pOneManager^.us_CoreSelect = usActiveCore then
      if pOneManager^.p_Functions <> NIL & pOneManager^.ud_CounterRt = ( aTaskInfoCore[usActiveCore].ud_MyRtTaskTime_us) then
        pOneManager^.p_Functions^.p_This^.UpdateRtPostscan();
      end_if;
    end_if;
    pOneManager += SIZEOF(t_OneVaranManager);
  end_for;

END_FUNCTION

#pragma warning(disable:73);
FUNCTION HwControl::CalcTimeMeasurementPreScan
  VAR_INPUT
    pHwControlTimes 	: ^t_HwControl_Times_SINGLE;
  END_VAR
#pragma warning(default:73);

#ifdef HWCONTROL_TIME_MEASUREMENT
  if ops.tAbsolute > HWCONTROL_TIME_MEASUREMENT_DELAY then

    if pHwControlTimes^.sRtPreScan_Help.bRestart then

      pHwControlTimes^.sRtPrescan_Total.ActTime         := 0;
      pHwControlTimes^.sRtPrescan_Total.AvgTime         := 0;
      pHwControlTimes^.sRtPrescan_Total.MinTime         := 16#FFFF;
      pHwControlTimes^.sRtPrescan_Total.MaxTime         := 0;

      pHwControlTimes^.sRtPrescan_FirstCallHW.ActTime   := 0;
      pHwControlTimes^.sRtPrescan_FirstCallHW.AvgTime   := 0;
      pHwControlTimes^.sRtPrescan_FirstCallHW.MinTime   := 16#FFFF;
      pHwControlTimes^.sRtPrescan_FirstCallHW.MaxTime   := 0;

      pHwControlTimes^.sRtPrescan_Varan.ActTime         := 0;
      pHwControlTimes^.sRtPrescan_Varan.AvgTime         := 0;
      pHwControlTimes^.sRtPrescan_Varan.MinTime         := 16#FFFF;
      pHwControlTimes^.sRtPrescan_Varan.MaxTime         := 0;

      pHwControlTimes^.sRtPrescan_Other.ActTime         := 0;
      pHwControlTimes^.sRtPrescan_Other.AvgTime         := 0;
      pHwControlTimes^.sRtPrescan_Other.MinTime         := 16#FFFF;
      pHwControlTimes^.sRtPrescan_Other.MaxTime         := 0;

      pHwControlTimes^.sRtPrescan_HwObjects.ActTime     := 0;
      pHwControlTimes^.sRtPrescan_HwObjects.AvgTime     := 0;
      pHwControlTimes^.sRtPrescan_HwObjects.MinTime     := 16#FFFF;
      pHwControlTimes^.sRtPrescan_HwObjects.MaxTime     := 0;

      pHwControlTimes^.sRtPreScan_Help.udCycleCnt       := 0;
      pHwControlTimes^.sRtPreScan_Help.bRestart         := FALSE;
      pHwControlTimes^.sRtPreScan_Help.bFinished        := FALSE;

    elsif pHwControlTimes^.sRtPreScan_Help.bFinished = FALSE then

      pHwControlTimes^.sRtPreScan_Help.udCycleCnt  += 1;

      //First Call Objects Min/Max
      //*****************************************************************************
      if pHwControlTimes^.sRtPrescan_FirstCallHW.ActTime > pHwControlTimes^.sRtPrescan_FirstCallHW.MaxTime then
        pHwControlTimes^.sRtPrescan_FirstCallHW.MaxTime := pHwControlTimes^.sRtPrescan_FirstCallHW.ActTime;

      elsif pHwControlTimes^.sRtPrescan_FirstCallHW.ActTime < pHwControlTimes^.sRtPrescan_FirstCallHW.MinTime then
        pHwControlTimes^.sRtPrescan_FirstCallHW.MinTime := pHwControlTimes^.sRtPrescan_FirstCallHW.ActTime;
      end_if;

      //VARAN Objects Min/Max
      //*****************************************************************************
      if pHwControlTimes^.sRtPrescan_Varan.ActTime > pHwControlTimes^.sRtPrescan_Varan.MaxTime then
        pHwControlTimes^.sRtPrescan_Varan.MaxTime := pHwControlTimes^.sRtPrescan_Varan.ActTime;

      elsif pHwControlTimes^.sRtPrescan_Varan.ActTime < pHwControlTimes^.sRtPrescan_Varan.MinTime then
        pHwControlTimes^.sRtPrescan_Varan.MinTime := pHwControlTimes^.sRtPrescan_Varan.ActTime;
      end_if;

      //HwControl-Login Objects Min/Max
      //*****************************************************************************
      if pHwControlTimes^.sRtPrescan_HwObjects.ActTime > pHwControlTimes^.sRtPrescan_HwObjects.MaxTime then
        pHwControlTimes^.sRtPrescan_HwObjects.MaxTime := pHwControlTimes^.sRtPrescan_HwObjects.ActTime;

      elsif pHwControlTimes^.sRtPrescan_HwObjects.ActTime < pHwControlTimes^.sRtPrescan_HwObjects.MinTime then
        pHwControlTimes^.sRtPrescan_HwObjects.MinTime := pHwControlTimes^.sRtPrescan_HwObjects.ActTime;
      end_if;

      //Other Objects Min/Max (DIAS Master and Special HW)
      //*****************************************************************************
      if pHwControlTimes^.sRtPrescan_Other.ActTime > pHwControlTimes^.sRtPrescan_Other.MaxTime then
        pHwControlTimes^.sRtPrescan_Other.MaxTime := pHwControlTimes^.sRtPrescan_Other.ActTime;

      elsif pHwControlTimes^.sRtPrescan_Other.ActTime < pHwControlTimes^.sRtPrescan_Other.MinTime then
        pHwControlTimes^.sRtPrescan_Other.MinTime := pHwControlTimes^.sRtPrescan_Other.ActTime;
      end_if;

      //Calculate Total amount of realtime
      //*****************************************************************************
      pHwControlTimes^.sRtPrescan_Total.ActTime := pHwControlTimes^.sRtPrescan_FirstCallHW.ActTime +
                                                   pHwControlTimes^.sRtPrescan_Varan.ActTime +
                                                   pHwControlTimes^.sRtPrescan_HwObjects.ActTime +
                                                   pHwControlTimes^.sRtPrescan_Other.ActTime;
      //Total Realtime Min/Max
      //*****************************************************************************
      if pHwControlTimes^.sRtPrescan_Total.ActTime > pHwControlTimes^.sRtPrescan_Total.MaxTime then
        pHwControlTimes^.sRtPrescan_Total.MaxTime := pHwControlTimes^.sRtPrescan_Total.ActTime;

      elsif pHwControlTimes^.sRtPrescan_Total.ActTime < pHwControlTimes^.sRtPrescan_Total.MinTime then
        pHwControlTimes^.sRtPrescan_Total.MinTime := pHwControlTimes^.sRtPrescan_Total.ActTime;
      end_if;

      pHwControlTimes^.sRtPrescan_FirstCallHW.AvgTime   += pHwControlTimes^.sRtPrescan_FirstCallHW.ActTime;
      pHwControlTimes^.sRtPrescan_Varan.AvgTime         += pHwControlTimes^.sRtPrescan_Varan.ActTime;
      pHwControlTimes^.sRtPrescan_HwObjects.AvgTime     += pHwControlTimes^.sRtPrescan_HwObjects.ActTime;
      pHwControlTimes^.sRtPrescan_Other.AvgTime         += pHwControlTimes^.sRtPrescan_Other.ActTime;
      pHwControlTimes^.sRtPrescan_Total.AvgTime         += pHwControlTimes^.sRtPrescan_Total.ActTime;

      //Finished measurement?
      if pHwControlTimes^.sRtPreScan_Help.udCycleCnt >= HWCONTROL_TIME_MEASUREMENT_CNT then

        pHwControlTimes^.sRtPrescan_FirstCallHW.AvgTime   /= HWCONTROL_TIME_MEASUREMENT_CNT;
        pHwControlTimes^.sRtPrescan_Varan.AvgTime         /= HWCONTROL_TIME_MEASUREMENT_CNT;
        pHwControlTimes^.sRtPrescan_HwObjects.AvgTime     /= HWCONTROL_TIME_MEASUREMENT_CNT;
        pHwControlTimes^.sRtPrescan_Other.AvgTime         /= HWCONTROL_TIME_MEASUREMENT_CNT;
        pHwControlTimes^.sRtPrescan_Total.AvgTime         /= HWCONTROL_TIME_MEASUREMENT_CNT;

        pHwControlTimes^.sRtPreScan_Help.bFinished         := TRUE;
      end_if;
    end_if;
  end_if;
#endif

END_FUNCTION

#pragma warning(disable:73);
FUNCTION HwControl::CalcTimeMeasurementPostScan
  VAR_INPUT
    pHwControlTimes 	: ^t_HwControl_Times_SINGLE;
  END_VAR
#pragma warning(default:73);

#ifdef HWCONTROL_TIME_MEASUREMENT
  if ops.tAbsolute > HWCONTROL_TIME_MEASUREMENT_DELAY then

    if pHwControlTimes^.sRtPostScan_Help.bRestart then

      pHwControlTimes^.sRtPostscan_Total.ActTime      := 0;
      pHwControlTimes^.sRtPostscan_Total.AvgTime      := 0;
      pHwControlTimes^.sRtPostscan_Total.MinTime      := 16#FFFF;
      pHwControlTimes^.sRtPostscan_Total.MaxTime      := 0;

      pHwControlTimes^.sRtPostscan_Varan.ActTime      := 0;
      pHwControlTimes^.sRtPostscan_Varan.AvgTime      := 0;
      pHwControlTimes^.sRtPostscan_Varan.MinTime      := 16#FFFF;
      pHwControlTimes^.sRtPostscan_Varan.MaxTime      := 0;

      pHwControlTimes^.sRtPostscan_HwObjects.ActTime  := 0;
      pHwControlTimes^.sRtPostscan_HwObjects.AvgTime  := 0;
      pHwControlTimes^.sRtPostscan_HwObjects.MinTime  := 16#FFFF;
      pHwControlTimes^.sRtPostscan_HwObjects.MaxTime  := 0;

      pHwControlTimes^.sRtPostScan_Help.udCycleCnt    := 0;
      pHwControlTimes^.sRtPostScan_Help.bRestart      := FALSE;
      pHwControlTimes^.sRtPostScan_Help.bFinished     := FALSE;

    elsif pHwControlTimes^.sRtPostScan_Help.bFinished = FALSE then

      pHwControlTimes^.sRtPostScan_Help.udCycleCnt  += 1;

      //VARAN Objects Min/Max
      if pHwControlTimes^.sRtPostscan_Varan.ActTime > pHwControlTimes^.sRtPostscan_Varan.MaxTime then
        pHwControlTimes^.sRtPostscan_Varan.MaxTime := pHwControlTimes^.sRtPostscan_Varan.ActTime;

      elsif pHwControlTimes^.sRtPostscan_Varan.ActTime < pHwControlTimes^.sRtPostscan_Varan.MinTime then
        pHwControlTimes^.sRtPostscan_Varan.MinTime := pHwControlTimes^.sRtPostscan_Varan.ActTime;
      end_if;

      //HwControl-Login Objects Min/Max
      if pHwControlTimes^.sRtPostscan_HwObjects.ActTime > pHwControlTimes^.sRtPostscan_HwObjects.MaxTime then
        pHwControlTimes^.sRtPostscan_HwObjects.MaxTime := pHwControlTimes^.sRtPostscan_HwObjects.ActTime;

      elsif pHwControlTimes^.sRtPostscan_HwObjects.ActTime < pHwControlTimes^.sRtPostscan_HwObjects.MinTime then
        pHwControlTimes^.sRtPostscan_HwObjects.MinTime := pHwControlTimes^.sRtPostscan_HwObjects.ActTime;
      end_if;

      //Calculate Total amount of realtime
      pHwControlTimes^.sRtPostscan_Total.ActTime := pHwControlTimes^.sRtPostscan_Varan.ActTime +
                                                    pHwControlTimes^.sRtPostscan_HwObjects.ActTime;
      //Total Realtime Min/Max
      if pHwControlTimes^.sRtPostscan_Total.ActTime > pHwControlTimes^.sRtPostscan_Total.MaxTime then
        pHwControlTimes^.sRtPostscan_Total.MaxTime := pHwControlTimes^.sRtPostscan_Total.ActTime;

      elsif pHwControlTimes^.sRtPostscan_Total.ActTime < pHwControlTimes^.sRtPostscan_Total.MinTime then
        pHwControlTimes^.sRtPostscan_Total.MinTime := pHwControlTimes^.sRtPostscan_Total.ActTime;
      end_if;

      pHwControlTimes^.sRtPostscan_Varan.AvgTime         += pHwControlTimes^.sRtPostscan_Varan.ActTime;
      pHwControlTimes^.sRtPostscan_HwObjects.AvgTime     += pHwControlTimes^.sRtPostscan_HwObjects.ActTime;
      pHwControlTimes^.sRtPostscan_Total.AvgTime         += pHwControlTimes^.sRtPostscan_Total.ActTime;

      //Finished measurement?
      if pHwControlTimes^.sRtPostScan_Help.udCycleCnt >= HWCONTROL_TIME_MEASUREMENT_CNT then

        pHwControlTimes^.sRtPostscan_Varan.AvgTime           /= HWCONTROL_TIME_MEASUREMENT_CNT;
        pHwControlTimes^.sRtPostscan_HwObjects.AvgTime       /= HWCONTROL_TIME_MEASUREMENT_CNT;
        pHwControlTimes^.sRtPostscan_Total.AvgTime           /= HWCONTROL_TIME_MEASUREMENT_CNT;

        pHwControlTimes^.sRtPostScan_Help.bFinished   := TRUE;
      end_if;
    end_if;
  end_if;
#endif

END_FUNCTION

#pragma warning(disable:73);
FUNCTION HwControl::CalcTimeMeasurementCyclic
  VAR_INPUT
    pHwControlTimes 	: ^t_HwControl_Times_SINGLE;
  END_VAR
#pragma warning(default:73);

#ifdef HWCONTROL_TIME_MEASUREMENT
  if ops.tAbsolute > HWCONTROL_TIME_MEASUREMENT_DELAY then

    if pHwControlTimes^.sCywork_Help.bRestart then

      pHwControlTimes^.sCyWork_Total.ActTime         := 0;
      pHwControlTimes^.sCyWork_Total.AvgTime         := 0;
      pHwControlTimes^.sCyWork_Total.MinTime         := 16#FFFF;
      pHwControlTimes^.sCyWork_Total.MaxTime         := 0;

      pHwControlTimes^.sCyWork_Varan.ActTime         := 0;
      pHwControlTimes^.sCyWork_Varan.AvgTime         := 0;
      pHwControlTimes^.sCyWork_Varan.MinTime         := 16#FFFF;
      pHwControlTimes^.sCyWork_Varan.MaxTime         := 0;

      pHwControlTimes^.sCyWork_HwObjects.ActTime     := 0;
      pHwControlTimes^.sCyWork_HwObjects.AvgTime     := 0;
      pHwControlTimes^.sCyWork_HwObjects.MinTime     := 16#FFFF;
      pHwControlTimes^.sCyWork_HwObjects.MaxTime     := 0;

      pHwControlTimes^.sCywork_Help.udCycleCnt       := 0;
      pHwControlTimes^.sCywork_Help.bRestart         := FALSE;
      pHwControlTimes^.sCywork_Help.bFinished        := FALSE;

    elsif pHwControlTimes^.sCywork_Help.bFinished = FALSE then

      pHwControlTimes^.sCywork_Help.udCycleCnt  += 1;

      //VARAN Objects Min/Max
      if pHwControlTimes^.sCyWork_Varan.ActTime > pHwControlTimes^.sCyWork_Varan.MaxTime then
        pHwControlTimes^.sCyWork_Varan.MaxTime := pHwControlTimes^.sCyWork_Varan.ActTime;

      elsif pHwControlTimes^.sCyWork_Varan.ActTime < pHwControlTimes^.sCyWork_Varan.MinTime then
        pHwControlTimes^.sCyWork_Varan.MinTime := pHwControlTimes^.sCyWork_Varan.ActTime;
      end_if;

      //HwControl-Login Objects Min/Max
      if pHwControlTimes^.sCyWork_HwObjects.ActTime > pHwControlTimes^.sCyWork_HwObjects.MaxTime then
        pHwControlTimes^.sCyWork_HwObjects.MaxTime := pHwControlTimes^.sCyWork_HwObjects.ActTime;

      elsif pHwControlTimes^.sCyWork_HwObjects.ActTime < pHwControlTimes^.sCyWork_HwObjects.MinTime then
        pHwControlTimes^.sCyWork_HwObjects.MinTime := pHwControlTimes^.sCyWork_HwObjects.ActTime;
      end_if;

      //Calculate Total amount of realtime
      pHwControlTimes^.sCyWork_Total.ActTime := pHwControlTimes^.sCyWork_Varan.ActTime +
                                                   pHwControlTimes^.sCyWork_HwObjects.ActTime;
      //Total Realtime Min/Max
      if pHwControlTimes^.sCyWork_Total.ActTime > pHwControlTimes^.sCyWork_Total.MaxTime then
        pHwControlTimes^.sCyWork_Total.MaxTime := pHwControlTimes^.sCyWork_Total.ActTime;

      elsif pHwControlTimes^.sCyWork_Total.ActTime < pHwControlTimes^.sCyWork_Total.MinTime then
        pHwControlTimes^.sCyWork_Total.MinTime := pHwControlTimes^.sCyWork_Total.ActTime;
      end_if;

      pHwControlTimes^.sCyWork_Varan.AvgTime         += pHwControlTimes^.sCyWork_Varan.ActTime;
      pHwControlTimes^.sCyWork_HwObjects.AvgTime     += pHwControlTimes^.sCyWork_HwObjects.ActTime;
      pHwControlTimes^.sCyWork_Total.AvgTime         += pHwControlTimes^.sCyWork_Total.ActTime;

      //Finished measurement?
      if pHwControlTimes^.sCywork_Help.udCycleCnt >= HWCONTROL_TIME_MEASUREMENT_CNT then

        pHwControlTimes^.sCyWork_Varan.AvgTime           /= HWCONTROL_TIME_MEASUREMENT_CNT;
        pHwControlTimes^.sCyWork_HwObjects.AvgTime       /= HWCONTROL_TIME_MEASUREMENT_CNT;
        pHwControlTimes^.sCyWork_Total.AvgTime           /= HWCONTROL_TIME_MEASUREMENT_CNT;

        pHwControlTimes^.sCywork_Help.bFinished   := TRUE;
      end_if;
    end_if;
  end_if;
#endif
END_FUNCTION

FUNCTION HwControl::UpdateRtFirstCallObjects
  VAR_INPUT
    usCoreSelect 	: USINT;
  END_VAR
  VAR
    pHelpCallFirst  : ^t_HwObjectListCallFirst;
  END_VAR

  // special classes with first call priority, which are controlled by HwControl
  if pCallFirstObjects then
    pHelpCallFirst := pCallFirstObjects;
    while pHelpCallFirst <> NIL do
      if pHelpCallFirst^.us_CoreSelect = usCoreSelect then
      pHelpCallFirst^.pThis^.RtWork(0);
      end_if;
      pHelpCallFirst := pHelpCallFirst^.pNext;
    end_while;
    // Record finish of first object call. p4 = "HwCo" as ascii (1.215.775.599 = 0x4857434F = "HwCo")
    OS_MakeTraceEntry(pSystrace, HWCONTROL_SYSTRACE_TYPE, HWCONTROL_SYSTRACE_RTPRESCAN_FINISHED_FIRST_CALL_OBJECTS, usCoreSelect);
  end_if;

END_FUNCTION

FUNCTION HwControl::UpdateRtLoginObjects
  VAR_INPUT
    usCoreSelect 	: USINT;
  END_VAR
  VAR
    pHelp           : ^t_HwObjectListElement;
  END_VAR

  // objects, which are controlled by HwControl
  if pHwControlLogins then
    pHelp := pHwControlLogins;
    while pHelp <> NIL do
      if pHelp^.bdSettings.RtPreScan & pHelp^.us_CoreSelect = usCoreSelect then
        pHelp^.pThis^.RtWork(CALL_OPTION_RT_PRESCAN);
      end_if;
      pHelp := pHelp^.pNext;
    end_while;
  end_if;

END_FUNCTION

FUNCTION HwControl::UpdateRtPostscanLoginObjects
  VAR_INPUT
    usCoreSelect 	: USINT;
  END_VAR
  VAR
    pHelp           : ^t_HwObjectListElement;
  END_VAR

  // objects, which are controlled by HwControl
  if pHwControlLogins then
    pHelp := pHwControlLogins;
    while pHelp <> NIL do
      if pHelp^.bdSettings.RtPostScan & pHelp^.us_CoreSelect = usCoreSelect then
        pHelp^.pThis^.RtWork(CALL_OPTION_RT_POSTSCAN);
      end_if;
      pHelp := pHelp^.pNext;
    end_while;
  end_if;

END_FUNCTION

FUNCTION HwControl::CalculateTaskInfo
  VAR_INPUT
    us_CoreSelect 	: USINT;
    pTaskInfo 	    : ^t_s_TaskCoreInfo;
  END_VAR
  VAR
    pHelp           : ^t_HwObjectListElement;
    pFirstCall      : ^t_HwObjectListCallFirst;
    pOneManager     : ^t_OneVaranManager;
    CurrGGT         : UDINT;
    i               : USINT;
  END_VAR

  //Calculate GGT of all objects (HwObjects, VaranManager, FirstCallHW and DiasMaster)

  //Calculate for Realtime
  //**************************************************************************************************************
  CurrGGT := 0;   //Start with 0

  //Go through all varanmanagers
  pOneManager := #a_VaranManager[0];
  for i := 0 to ( MAX_VARAN_MANAGERS - 1 ) do

    //Check if manager is available, set for right core and has set a time
    if ( pOneManager^.p_Functions         <> NIL
       & pOneManager^.p_Functions^.p_This <> NIL
       & pOneManager^.ud_RtTime_us        <> 0
       & pOneManager^.us_CoreSelect        = us_CoreSelect
       )
    then
      CurrGGT := CalculateGGT(Var1:=CurrGGT, Var2:=pOneManager^.ud_RtTime_us);
    end_if;
    pOneManager += sizeof(t_OneVaranManager);
  end_for;

  pHelp := pHwControlLogins;

  //Go through all HwObjects
  while pHelp <> NIL do
    if pHelp^.ud_RtTime_us & pHelp^.us_CoreSelect = us_CoreSelect then
      CurrGGT := CalculateGGT(Var1:=CurrGGT, Var2:=pHelp^.ud_RtTime_us);
    end_if;
    pHelp := pHelp^.pNext;
  end_while;

  pFirstCall := pCallFirstObjects;

  //Go through all first call objects
  while pFirstCall <> NIL do
    if pFirstCall^.ud_RtTime_us & pFirstCall^.us_CoreSelect = us_CoreSelect then
      CurrGGT := CalculateGGT(Var1:=CurrGGT, Var2:=pFirstCall^.ud_RtTime_us);
    end_if;
    pFirstCall := pFirstCall^.pNext;
  end_while;

  //Also calculate with DIAS Master time (DIAS only runs on core 0)
  if us_CoreSelect = TASK_SELECT_CORE0 then
    if s_DiasMaster.p_Functions <> NIL & s_DiasMaster.p_Functions^.ud_DiasTime then
      CurrGGT := CalculateGGT(Var1:=CurrGGT, Var2:=s_DiasMaster.p_Functions^.ud_DiasTime);
    end_if;
  end_if;

  //Core 0: set to maintimer if no one wants a time
  if ( us_CoreSelect = TASK_SELECT_CORE0 ) & ( CurrGGT = 0 ) then
    CurrGGT := _Clockticks;
  end_if;

  //Check if maintimer is fast enough
  if ( CurrGGT <> 0 ) & ( CurrGGT < _ClockTicks ) then
    HWC_LogValue2(this,"@0179 (HwControl::CalculateTaskInfo) Calc RtTaskTime: Maintimersetting is too slow. Needed maintimer: 0x{0} µs, Actual Maintimer: 0x{1} µs", CurrGGT,_ClockTicks);
    HwControl::State := _InvalidConfguration;
    return;
  end_if;

  //Save realtime task time
  pTaskInfo^.ud_MyRtTaskTime_us := CurrGGT;

  //Calculate for Cyclic
  //**************************************************************************************************************
  CurrGGT := 0; //Start with 0

  //Go through all varanmanagers
  pOneManager := #a_VaranManager[0];
  for i := 0 to ( MAX_VARAN_MANAGERS - 1 ) do

    //Check if manager is available, set for right core and has set a time
    if ( pOneManager^.p_Functions         <> NIL
       & pOneManager^.p_Functions^.p_This <> NIL
       & pOneManager^.ud_CyTime_us        <> 0
       & pOneManager^.us_CoreSelect        = us_CoreSelect
       )
    then
      CurrGGT := CalculateGGT(Var1:=CurrGGT, Var2:=pOneManager^.ud_CyTime_us);
    end_if;

    pOneManager += sizeof(t_OneVaranManager);
  end_for;

  pHelp := pHwControlLogins;

  //Go through all HwObjects
  while pHelp <> NIL do
    if pHelp^.ud_CyTime_us & pHelp^.us_CoreSelect = us_CoreSelect then
      CurrGGT := CalculateGGT(Var1:=CurrGGT, Var2:=pHelp^.ud_CyTime_us);
    end_if;
    pHelp := pHelp^.pNext;
  end_while;

  pFirstCall := pCallFirstObjects;

  //Go through all first call objects
  while pFirstCall <> NIL do
    if pFirstCall^.ud_CyTime_us & pFirstCall^.us_CoreSelect = us_CoreSelect then
      CurrGGT := CalculateGGT(Var1:=CurrGGT, Var2:=pFirstCall^.ud_CyTime_us);
    end_if;
    pFirstCall := pFirstCall^.pNext;
  end_while;

  //Core 0: set to maintimer if no one wants a time
  if ( us_CoreSelect = TASK_SELECT_CORE0 ) & ( CurrGGT = 0 ) then
    CurrGGT := _Clockticks;
  end_if;

  //Check if maintimer is fast enough
  if ( CurrGGT <> 0 ) & ( CurrGGT < _ClockTicks ) then
    HWC_LogValue2(this,"@017A (HwControl::CalculateTaskInfo) Calc CyTaskTime: Maintimersetting is too slow. Needed maintimer: 0x{0} µs, Actual Maintimer: 0x{1} µs", CurrGGT,_ClockTicks);
    HwControl::State := _InvalidConfguration;
    return;
  end_if;

  //Save realtime task time
  pTaskInfo^.ud_MyCyTaskTime_us := CurrGGT;

END_FUNCTION

FUNCTION HwControl::CalculateGGT
  VAR_INPUT
    Var1 	: UDINT;
    Var2 	: UDINT;
  END_VAR
  VAR_OUTPUT
    ggT 	: UDINT;
  END_VAR

  if Var2 = 0 then
    ggT := Var1;
  else
    ggT := CalculateGGT(Var1:=Var2, Var2:=Var1 MOD Var2);
  end_if;

END_FUNCTION

FUNCTION HwControl::Get_ITASK_Version
  VAR_OUTPUT
    version 	: UDINT;
  END_VAR

  // Anm.: Beim Salamander darf das udVersion Element aus der LSL_ITASK Struktur
  // (Makro OS_ITASK_VERSION) erst ab 09.03.080 interpretiert werden, weil sonst
  // keine Versionsnummer dahintersteckt, sondern ein Funktionszeiger auf eine Dummy-Funktion.
  // Die Versionen im Salamander, bei denen udVersion gültig ist:
  //  9.3 er Versionen:   ab 09.03.080
  //  9.2 er Versionen:   ab 09.02.049

  IF _RtOSVersion < 16#9000 | _RtOSVersion >= 16#9350 THEN
    version := OS_ITASK_VERSION;
  ELSIF _RtOSVersion < 16#9300 & _RtOSVersion >= 16#9231 THEN
    version := OS_ITASK_VERSION;
  ELSE
    version := 0;
  END_IF;

END_FUNCTION

FUNCTION VIRTUAL GLOBAL HwControl::UpdateRtPostScan
VAR
  us_CoreSelect : USINT;
END_VAR

  us_CoreSelect := TASK_SELECT_CORE0;
  RtPostScan_CoreX(pCoreSelect:=#us_CoreSelect);

END_FUNCTION

FUNCTION VIRTUAL GLOBAL HwControl::CyWork
  VAR_INPUT
    EAX 	: UDINT;
  END_VAR
  VAR_OUTPUT
    state (EAX) 	: UDINT;
  END_VAR
  VAR
    us_CoreSelect : USINT;
  END_VAR

  us_CoreSelect := TASK_SELECT_CORE0;
  CyWork_CoreX(pCoreSelect:=#us_CoreSelect);

  state := READY;

END_FUNCTION

FUNCTION GLOBAL __cdecl HWC_ops_cpuequipment_get
VAR_OUTPUT
  retcode : UDINT;
END_VAR
VAR
  ptr : ^UDINT;
END_VAR
  // we take the offset from _RealMaximumTime because an define for the right address would make troubles
  ptr := #_RealMaximumTime;
  ptr += 16#F44;
  retcode := ptr^;
END_FUNCTION

FUNCTION GLOBAL __cdecl HWC_ops_platform_get
VAR_OUTPUT
  retcode : UDINT;
END_VAR
  retcode := HWC_ops_cpuequipment_get() AND HWCONTROL_OPS_PLATFORMMASK;
END_FUNCTION

FUNCTION GLOBAL __cdecl HWC_ops_is_linux
VAR_OUTPUT
  retcode : UDINT;
END_VAR
  retcode := (HWC_ops_cpuequipment_get() AND (HWCONTROL_OPS_OS_LINUX OR HWCONTROL_OPS_EQUIPMENT_VALID)) = (HWCONTROL_OPS_OS_LINUX OR HWCONTROL_OPS_EQUIPMENT_VALID);
END_FUNCTION

FUNCTION GLOBAL __cdecl HWC_ops_is_salamander
VAR_OUTPUT
  retcode : UDINT;
END_VAR
  // wenn es ein Linux ist und platform = LSL_LASALOS dann ist es auch ein Salamander
  // bei platform = LSL_SALAMANDER ist es Salamander
  if HWC_ops_is_linux() &
    (HWC_ops_platform_get() = HWCONTROL_OPS_LASALOS |
     HWC_ops_platform_get() = HWCONTROL_OPS_SALAMANDER) then
    retcode := 1;
  else
    retcode := 0;
  end_if;
END_FUNCTION

FUNCTION GLOBAL __cdecl HWC_ops_is_gecko
VAR_OUTPUT
  retcode :UDINT;
END_VAR
  if HWC_ops_is_linux() &
    (HWC_ops_platform_get() = HWCONTROL_OPS_GECKO) then
    retcode := 1;
  else
    retcode := 0;
  end_if;
END_FUNCTION

FUNCTION GLOBAL __cdecl HWC_IsPostInitFinished
VAR_OUTPUT
  retcode : BOOL;
END_VAR

  retcode := bPostInitFinished;

END_FUNCTION
